(* IEC 61131-3 sources: plc-iiot-stack/flagship/src/POUs/Iiot/FB_IiotKnsMap, 8 files *)

(* ---- ApplyCommand.method.decl.st ---- *)
// Записать принятую команду строки diRule белого списка в GVL_Hmi или GVL_Station (импульс или rValue).
METHOD ApplyCommand : BOOL
VAR_INPUT
    diRule : DINT;
    rValue : REAL;
END_VAR

(* ---- ApplyCommand.method.impl.st ---- *)
ApplyCommand := TRUE;
CASE diRule OF
    1:  // P101 SetAuto
        GVL_Hmi.stP101Cmd.stCommon.xSetAuto := TRUE;
    2:  // P101 SetManual
        GVL_Hmi.stP101Cmd.stCommon.xSetManual := TRUE;
    3:  // P101 Start
        GVL_Hmi.stP101Cmd.xStart := TRUE;
    4:  // P101 Stop
        GVL_Hmi.stP101Cmd.xStop := TRUE;
    5:  // P101 SpeedSp
        GVL_Hmi.stP101Cmd.rSpeedSp_pct := rValue;
    6:  // P101 Ack
        GVL_Hmi.stP101Cmd.stCommon.xAck := TRUE;
    7:  // P101 Reset
        GVL_Hmi.stP101Cmd.stCommon.xReset := TRUE;
    8:  // P102 SetAuto
        GVL_Hmi.stP102Cmd.stCommon.xSetAuto := TRUE;
    9:  // P102 SetManual
        GVL_Hmi.stP102Cmd.stCommon.xSetManual := TRUE;
    10:  // P102 Start
        GVL_Hmi.stP102Cmd.xStart := TRUE;
    11:  // P102 Stop
        GVL_Hmi.stP102Cmd.xStop := TRUE;
    12:  // P102 SpeedSp
        GVL_Hmi.stP102Cmd.rSpeedSp_pct := rValue;
    13:  // P102 Ack
        GVL_Hmi.stP102Cmd.stCommon.xAck := TRUE;
    14:  // P102 Reset
        GVL_Hmi.stP102Cmd.stCommon.xReset := TRUE;
    15:  // P103 SetAuto
        GVL_Hmi.stP103Cmd.stCommon.xSetAuto := TRUE;
    16:  // P103 SetManual
        GVL_Hmi.stP103Cmd.stCommon.xSetManual := TRUE;
    17:  // P103 Start
        GVL_Hmi.stP103Cmd.xStart := TRUE;
    18:  // P103 Stop
        GVL_Hmi.stP103Cmd.xStop := TRUE;
    19:  // P103 SpeedSp
        GVL_Hmi.stP103Cmd.rSpeedSp_pct := rValue;
    20:  // P103 Ack
        GVL_Hmi.stP103Cmd.stCommon.xAck := TRUE;
    21:  // P103 Reset
        GVL_Hmi.stP103Cmd.stCommon.xReset := TRUE;
    22:  // V1 SetAuto
        GVL_Hmi.stV1Cmd.stCommon.xSetAuto := TRUE;
    23:  // V1 SetManual
        GVL_Hmi.stV1Cmd.stCommon.xSetManual := TRUE;
    24:  // V1 Start
        GVL_Hmi.stV1Cmd.xStart := TRUE;
    25:  // V1 Stop
        GVL_Hmi.stV1Cmd.xStop := TRUE;
    26:  // V1 Ack
        GVL_Hmi.stV1Cmd.stCommon.xAck := TRUE;
    27:  // V1 Reset
        GVL_Hmi.stV1Cmd.stCommon.xReset := TRUE;
    28:  // LT101 Ack
        GVL_Hmi.stLT101Cmd.stCommon.xAck := TRUE;
    29:  // LT101 Reset
        GVL_Hmi.stLT101Cmd.stCommon.xReset := TRUE;
    30:  // LS102 Ack
        GVL_Hmi.stLS102Cmd.stCommon.xAck := TRUE;
    31:  // LS102 Reset
        GVL_Hmi.stLS102Cmd.stCommon.xReset := TRUE;
    32:  // LS103 Ack
        GVL_Hmi.stLS103Cmd.stCommon.xAck := TRUE;
    33:  // LS103 Reset
        GVL_Hmi.stLS103Cmd.stCommon.xReset := TRUE;
    34:  // IT111 Ack
        GVL_Hmi.stIT111Cmd.stCommon.xAck := TRUE;
    35:  // IT111 Reset
        GVL_Hmi.stIT111Cmd.stCommon.xReset := TRUE;
    36:  // TS112 Ack
        GVL_Hmi.stTS112Cmd.stCommon.xAck := TRUE;
    37:  // TS112 Reset
        GVL_Hmi.stTS112Cmd.stCommon.xReset := TRUE;
    38:  // MS113 Ack
        GVL_Hmi.stMS113Cmd.stCommon.xAck := TRUE;
    39:  // MS113 Reset
        GVL_Hmi.stMS113Cmd.stCommon.xReset := TRUE;
    40:  // IT121 Ack
        GVL_Hmi.stIT121Cmd.stCommon.xAck := TRUE;
    41:  // IT121 Reset
        GVL_Hmi.stIT121Cmd.stCommon.xReset := TRUE;
    42:  // TS122 Ack
        GVL_Hmi.stTS122Cmd.stCommon.xAck := TRUE;
    43:  // TS122 Reset
        GVL_Hmi.stTS122Cmd.stCommon.xReset := TRUE;
    44:  // MS123 Ack
        GVL_Hmi.stMS123Cmd.stCommon.xAck := TRUE;
    45:  // MS123 Reset
        GVL_Hmi.stMS123Cmd.stCommon.xReset := TRUE;
    46:  // IT131 Ack
        GVL_Hmi.stIT131Cmd.stCommon.xAck := TRUE;
    47:  // IT131 Reset
        GVL_Hmi.stIT131Cmd.stCommon.xReset := TRUE;
    48:  // TS132 Ack
        GVL_Hmi.stTS132Cmd.stCommon.xAck := TRUE;
    49:  // TS132 Reset
        GVL_Hmi.stTS132Cmd.stCommon.xReset := TRUE;
    50:  // MS133 Ack
        GVL_Hmi.stMS133Cmd.stCommon.xAck := TRUE;
    51:  // MS133 Reset
        GVL_Hmi.stMS133Cmd.stCommon.xReset := TRUE;
    52:  // PT201 Ack
        GVL_Hmi.stPT201Cmd.stCommon.xAck := TRUE;
    53:  // PT201 Reset
        GVL_Hmi.stPT201Cmd.stCommon.xReset := TRUE;
    54:  // FT202 Ack
        GVL_Hmi.stFT202Cmd.stCommon.xAck := TRUE;
    55:  // FT202 Reset
        GVL_Hmi.stFT202Cmd.stCommon.xReset := TRUE;
    56:  // LS203 Ack
        GVL_Hmi.stLS203Cmd.stCommon.xAck := TRUE;
    57:  // LS203 Reset
        GVL_Hmi.stLS203Cmd.stCommon.xReset := TRUE;
    58:  // ES301 Ack
        GVL_Hmi.stES301Cmd.stCommon.xAck := TRUE;
    59:  // ES301 Reset
        GVL_Hmi.stES301Cmd.stCommon.xReset := TRUE;
    60:  // YS302 Ack
        GVL_Hmi.stYS302Cmd.stCommon.xAck := TRUE;
    61:  // YS302 Reset
        GVL_Hmi.stYS302Cmd.stCommon.xReset := TRUE;
    62:  // YS303 Ack
        GVL_Hmi.stYS303Cmd.stCommon.xAck := TRUE;
    63:  // YS303 Reset
        GVL_Hmi.stYS303Cmd.stCommon.xReset := TRUE;
    64:  // AT401 Ack
        GVL_Hmi.stAT401Cmd.stCommon.xAck := TRUE;
    65:  // AT401 Reset
        GVL_Hmi.stAT401Cmd.stCommon.xReset := TRUE;
    66:  // AT402 Ack
        GVL_Hmi.stAT402Cmd.stCommon.xAck := TRUE;
    67:  // AT402 Reset
        GVL_Hmi.stAT402Cmd.stCommon.xReset := TRUE;
    68:  // TT403 Ack
        GVL_Hmi.stTT403Cmd.stCommon.xAck := TRUE;
    69:  // TT403 Reset
        GVL_Hmi.stTT403Cmd.stCommon.xReset := TRUE;
    70:  // ZS404 Ack
        GVL_Hmi.stZS404Cmd.stCommon.xAck := TRUE;
    71:  // ZS404 Reset
        GVL_Hmi.stZS404Cmd.stCommon.xReset := TRUE;
    72:  // YS405 Ack
        GVL_Hmi.stYS405Cmd.stCommon.xAck := TRUE;
    73:  // YS405 Reset
        GVL_Hmi.stYS405Cmd.stCommon.xReset := TRUE;
    74:  // HS501 Ack
        GVL_Hmi.stHS501Cmd.stCommon.xAck := TRUE;
    75:  // HS501 Reset
        GVL_Hmi.stHS501Cmd.stCommon.xReset := TRUE;
    76:  // HS502 Ack
        GVL_Hmi.stHS502Cmd.stCommon.xAck := TRUE;
    77:  // HS502 Reset
        GVL_Hmi.stHS502Cmd.stCommon.xReset := TRUE;
    78:  // KNS1 SetAuto
        GVL_Station.stStationCmd.xSetAuto := TRUE;
    79:  // KNS1 SetManual
        GVL_Station.stStationCmd.xSetManual := TRUE;
    80:  // KNS1 SetStepped
        GVL_Station.stStationCmd.xSetStepped := TRUE;
    81:  // KNS1 SetLevelPid
        GVL_Station.stStationCmd.xSetLevelPid := TRUE;
    82:  // KNS1 AckAll
        GVL_Station.stStationCmd.xAckAll := TRUE;
    83:  // KNS1 ResetAll
        GVL_Station.stStationCmd.xResetAll := TRUE;
    84:  // KNS1 Silence
        GVL_Station.stStationCmd.xSilence := TRUE;
    85:  // LIC101 SetAuto
        GVL_Station.stLIC101Cmd.stCommon.xSetAuto := TRUE;
    86:  // LIC101 SetManual
        GVL_Station.stLIC101Cmd.stCommon.xSetManual := TRUE;
ELSE
    ApplyCommand := FALSE;
END_CASE

(* ---- DeviceCmdState.method.decl.st ---- *)
// Счётчик обработанных команд и результат последней команды устройства diDev (ST_IiotCmdRule.diDev).
METHOD DeviceCmdState
VAR_INPUT
    diDev : DINT;
END_VAR
VAR_OUTPUT
    uiSeq : UINT;
    iResult : INT;
END_VAR

(* ---- DeviceCmdState.method.impl.st ---- *)
uiSeq := 0;
iResult := 0;
CASE diDev OF
    1:  // P101
        uiSeq := GVL_Devices.fbP101.stSts.stCommon.uiCmdSeq;
        iResult := TO_INT(GVL_Devices.fbP101.stSts.stCommon.eCmdResult);
    2:  // P102
        uiSeq := GVL_Devices.fbP102.stSts.stCommon.uiCmdSeq;
        iResult := TO_INT(GVL_Devices.fbP102.stSts.stCommon.eCmdResult);
    3:  // P103
        uiSeq := GVL_Devices.fbP103.stSts.stCommon.uiCmdSeq;
        iResult := TO_INT(GVL_Devices.fbP103.stSts.stCommon.eCmdResult);
    4:  // V1
        uiSeq := GVL_Devices.fbV1.stSts.stCommon.uiCmdSeq;
        iResult := TO_INT(GVL_Devices.fbV1.stSts.stCommon.eCmdResult);
    5:  // LT101
        uiSeq := GVL_Devices.fbLT101.stSts.stCommon.uiCmdSeq;
        iResult := TO_INT(GVL_Devices.fbLT101.stSts.stCommon.eCmdResult);
    6:  // LS102
        uiSeq := GVL_Devices.fbLS102.stSts.stCommon.uiCmdSeq;
        iResult := TO_INT(GVL_Devices.fbLS102.stSts.stCommon.eCmdResult);
    7:  // LS103
        uiSeq := GVL_Devices.fbLS103.stSts.stCommon.uiCmdSeq;
        iResult := TO_INT(GVL_Devices.fbLS103.stSts.stCommon.eCmdResult);
    8:  // IT111
        uiSeq := GVL_Devices.fbIT111.stSts.stCommon.uiCmdSeq;
        iResult := TO_INT(GVL_Devices.fbIT111.stSts.stCommon.eCmdResult);
    9:  // TS112
        uiSeq := GVL_Devices.fbTS112.stSts.stCommon.uiCmdSeq;
        iResult := TO_INT(GVL_Devices.fbTS112.stSts.stCommon.eCmdResult);
    10:  // MS113
        uiSeq := GVL_Devices.fbMS113.stSts.stCommon.uiCmdSeq;
        iResult := TO_INT(GVL_Devices.fbMS113.stSts.stCommon.eCmdResult);
    11:  // IT121
        uiSeq := GVL_Devices.fbIT121.stSts.stCommon.uiCmdSeq;
        iResult := TO_INT(GVL_Devices.fbIT121.stSts.stCommon.eCmdResult);
    12:  // TS122
        uiSeq := GVL_Devices.fbTS122.stSts.stCommon.uiCmdSeq;
        iResult := TO_INT(GVL_Devices.fbTS122.stSts.stCommon.eCmdResult);
    13:  // MS123
        uiSeq := GVL_Devices.fbMS123.stSts.stCommon.uiCmdSeq;
        iResult := TO_INT(GVL_Devices.fbMS123.stSts.stCommon.eCmdResult);
    14:  // IT131
        uiSeq := GVL_Devices.fbIT131.stSts.stCommon.uiCmdSeq;
        iResult := TO_INT(GVL_Devices.fbIT131.stSts.stCommon.eCmdResult);
    15:  // TS132
        uiSeq := GVL_Devices.fbTS132.stSts.stCommon.uiCmdSeq;
        iResult := TO_INT(GVL_Devices.fbTS132.stSts.stCommon.eCmdResult);
    16:  // MS133
        uiSeq := GVL_Devices.fbMS133.stSts.stCommon.uiCmdSeq;
        iResult := TO_INT(GVL_Devices.fbMS133.stSts.stCommon.eCmdResult);
    17:  // PT201
        uiSeq := GVL_Devices.fbPT201.stSts.stCommon.uiCmdSeq;
        iResult := TO_INT(GVL_Devices.fbPT201.stSts.stCommon.eCmdResult);
    18:  // FT202
        uiSeq := GVL_Devices.fbFT202.stSts.stCommon.uiCmdSeq;
        iResult := TO_INT(GVL_Devices.fbFT202.stSts.stCommon.eCmdResult);
    19:  // LS203
        uiSeq := GVL_Devices.fbLS203.stSts.stCommon.uiCmdSeq;
        iResult := TO_INT(GVL_Devices.fbLS203.stSts.stCommon.eCmdResult);
    20:  // ES301
        uiSeq := GVL_Devices.fbES301.stSts.stCommon.uiCmdSeq;
        iResult := TO_INT(GVL_Devices.fbES301.stSts.stCommon.eCmdResult);
    21:  // YS302
        uiSeq := GVL_Devices.fbYS302.stSts.stCommon.uiCmdSeq;
        iResult := TO_INT(GVL_Devices.fbYS302.stSts.stCommon.eCmdResult);
    22:  // YS303
        uiSeq := GVL_Devices.fbYS303.stSts.stCommon.uiCmdSeq;
        iResult := TO_INT(GVL_Devices.fbYS303.stSts.stCommon.eCmdResult);
    23:  // AT401
        uiSeq := GVL_Devices.fbAT401.stSts.stCommon.uiCmdSeq;
        iResult := TO_INT(GVL_Devices.fbAT401.stSts.stCommon.eCmdResult);
    24:  // AT402
        uiSeq := GVL_Devices.fbAT402.stSts.stCommon.uiCmdSeq;
        iResult := TO_INT(GVL_Devices.fbAT402.stSts.stCommon.eCmdResult);
    25:  // TT403
        uiSeq := GVL_Devices.fbTT403.stSts.stCommon.uiCmdSeq;
        iResult := TO_INT(GVL_Devices.fbTT403.stSts.stCommon.eCmdResult);
    26:  // ZS404
        uiSeq := GVL_Devices.fbZS404.stSts.stCommon.uiCmdSeq;
        iResult := TO_INT(GVL_Devices.fbZS404.stSts.stCommon.eCmdResult);
    27:  // YS405
        uiSeq := GVL_Devices.fbYS405.stSts.stCommon.uiCmdSeq;
        iResult := TO_INT(GVL_Devices.fbYS405.stSts.stCommon.eCmdResult);
    28:  // HS501
        uiSeq := GVL_Devices.fbHS501.stSts.stCommon.uiCmdSeq;
        iResult := TO_INT(GVL_Devices.fbHS501.stSts.stCommon.eCmdResult);
    29:  // HS502
        uiSeq := GVL_Devices.fbHS502.stSts.stCommon.uiCmdSeq;
        iResult := TO_INT(GVL_Devices.fbHS502.stSts.stCommon.eCmdResult);
    30:  // KNS1
        uiSeq := GVL_Station.stStationSts.uiCmdSeq;
        iResult := TO_INT(GVL_Station.stStationSts.eCmdResult);
    31:  // LIC101
        uiSeq := GVL_Station.fbLIC101.stSts.stCommon.uiCmdSeq;
        iResult := TO_INT(GVL_Station.fbLIC101.stSts.stCommon.eCmdResult);
END_CASE

(* ---- FillAlarmWords.method.decl.st ---- *)
// Слова тревог устройств и станции (строки — источники перечня тревог по порядку ALARM_CFG.diWords).
METHOD FillAlarmWords
VAR_IN_OUT
    aWordTable : ARRAY[*] OF ST_IiotAlarmWords;
END_VAR

(* ---- FillAlarmWords.method.impl.st ---- *)
// Массив меньше перечня (не тот, что объявлен в PRG_Iiot): ничего не пишем, а не выходим за границы
IF LOWER_BOUND(aWordTable, 1) > 1 OR UPPER_BOUND(aWordTable, 1) < GVL_IiotMap.ALARM_WORDS_COUNT THEN
    RETURN;
END_IF
aWordTable[1].wActive := GVL_Devices.fbP101.stSts.stCommon.wAlmActive;
aWordTable[1].wUnack := GVL_Devices.fbP101.stSts.stCommon.wAlmUnack;
aWordTable[1].wShelved := GVL_Devices.fbP101.stSts.stCommon.wAlmShelved;
aWordTable[1].wSuppressed := GVL_Devices.fbP101.stSts.stCommon.wAlmSuppressed;
aWordTable[1].xOutOfService := GVL_Devices.fbP101.stSts.stCommon.eMode = PL.E_DeviceMode.OutOfService;
aWordTable[2].wActive := GVL_Devices.fbP102.stSts.stCommon.wAlmActive;
aWordTable[2].wUnack := GVL_Devices.fbP102.stSts.stCommon.wAlmUnack;
aWordTable[2].wShelved := GVL_Devices.fbP102.stSts.stCommon.wAlmShelved;
aWordTable[2].wSuppressed := GVL_Devices.fbP102.stSts.stCommon.wAlmSuppressed;
aWordTable[2].xOutOfService := GVL_Devices.fbP102.stSts.stCommon.eMode = PL.E_DeviceMode.OutOfService;
aWordTable[3].wActive := GVL_Devices.fbP103.stSts.stCommon.wAlmActive;
aWordTable[3].wUnack := GVL_Devices.fbP103.stSts.stCommon.wAlmUnack;
aWordTable[3].wShelved := GVL_Devices.fbP103.stSts.stCommon.wAlmShelved;
aWordTable[3].wSuppressed := GVL_Devices.fbP103.stSts.stCommon.wAlmSuppressed;
aWordTable[3].xOutOfService := GVL_Devices.fbP103.stSts.stCommon.eMode = PL.E_DeviceMode.OutOfService;
aWordTable[4].wActive := GVL_Devices.fbV1.stSts.stCommon.wAlmActive;
aWordTable[4].wUnack := GVL_Devices.fbV1.stSts.stCommon.wAlmUnack;
aWordTable[4].wShelved := GVL_Devices.fbV1.stSts.stCommon.wAlmShelved;
aWordTable[4].wSuppressed := GVL_Devices.fbV1.stSts.stCommon.wAlmSuppressed;
aWordTable[4].xOutOfService := GVL_Devices.fbV1.stSts.stCommon.eMode = PL.E_DeviceMode.OutOfService;
aWordTable[5].wActive := GVL_Devices.fbLT101.stSts.stCommon.wAlmActive;
aWordTable[5].wUnack := GVL_Devices.fbLT101.stSts.stCommon.wAlmUnack;
aWordTable[5].wShelved := GVL_Devices.fbLT101.stSts.stCommon.wAlmShelved;
aWordTable[5].wSuppressed := GVL_Devices.fbLT101.stSts.stCommon.wAlmSuppressed;
aWordTable[5].xOutOfService := GVL_Devices.fbLT101.stSts.stCommon.eMode = PL.E_DeviceMode.OutOfService;
aWordTable[6].wActive := GVL_Devices.fbLS102.stSts.stCommon.wAlmActive;
aWordTable[6].wUnack := GVL_Devices.fbLS102.stSts.stCommon.wAlmUnack;
aWordTable[6].wShelved := GVL_Devices.fbLS102.stSts.stCommon.wAlmShelved;
aWordTable[6].wSuppressed := GVL_Devices.fbLS102.stSts.stCommon.wAlmSuppressed;
aWordTable[6].xOutOfService := GVL_Devices.fbLS102.stSts.stCommon.eMode = PL.E_DeviceMode.OutOfService;
aWordTable[7].wActive := GVL_Devices.fbLS103.stSts.stCommon.wAlmActive;
aWordTable[7].wUnack := GVL_Devices.fbLS103.stSts.stCommon.wAlmUnack;
aWordTable[7].wShelved := GVL_Devices.fbLS103.stSts.stCommon.wAlmShelved;
aWordTable[7].wSuppressed := GVL_Devices.fbLS103.stSts.stCommon.wAlmSuppressed;
aWordTable[7].xOutOfService := GVL_Devices.fbLS103.stSts.stCommon.eMode = PL.E_DeviceMode.OutOfService;
aWordTable[8].wActive := GVL_Devices.fbIT111.stSts.stCommon.wAlmActive;
aWordTable[8].wUnack := GVL_Devices.fbIT111.stSts.stCommon.wAlmUnack;
aWordTable[8].wShelved := GVL_Devices.fbIT111.stSts.stCommon.wAlmShelved;
aWordTable[8].wSuppressed := GVL_Devices.fbIT111.stSts.stCommon.wAlmSuppressed;
aWordTable[8].xOutOfService := GVL_Devices.fbIT111.stSts.stCommon.eMode = PL.E_DeviceMode.OutOfService;
aWordTable[9].wActive := GVL_Devices.fbTS112.stSts.stCommon.wAlmActive;
aWordTable[9].wUnack := GVL_Devices.fbTS112.stSts.stCommon.wAlmUnack;
aWordTable[9].wShelved := GVL_Devices.fbTS112.stSts.stCommon.wAlmShelved;
aWordTable[9].wSuppressed := GVL_Devices.fbTS112.stSts.stCommon.wAlmSuppressed;
aWordTable[9].xOutOfService := GVL_Devices.fbTS112.stSts.stCommon.eMode = PL.E_DeviceMode.OutOfService;
aWordTable[10].wActive := GVL_Devices.fbMS113.stSts.stCommon.wAlmActive;
aWordTable[10].wUnack := GVL_Devices.fbMS113.stSts.stCommon.wAlmUnack;
aWordTable[10].wShelved := GVL_Devices.fbMS113.stSts.stCommon.wAlmShelved;
aWordTable[10].wSuppressed := GVL_Devices.fbMS113.stSts.stCommon.wAlmSuppressed;
aWordTable[10].xOutOfService := GVL_Devices.fbMS113.stSts.stCommon.eMode = PL.E_DeviceMode.OutOfService;
aWordTable[11].wActive := GVL_Devices.fbIT121.stSts.stCommon.wAlmActive;
aWordTable[11].wUnack := GVL_Devices.fbIT121.stSts.stCommon.wAlmUnack;
aWordTable[11].wShelved := GVL_Devices.fbIT121.stSts.stCommon.wAlmShelved;
aWordTable[11].wSuppressed := GVL_Devices.fbIT121.stSts.stCommon.wAlmSuppressed;
aWordTable[11].xOutOfService := GVL_Devices.fbIT121.stSts.stCommon.eMode = PL.E_DeviceMode.OutOfService;
aWordTable[12].wActive := GVL_Devices.fbTS122.stSts.stCommon.wAlmActive;
aWordTable[12].wUnack := GVL_Devices.fbTS122.stSts.stCommon.wAlmUnack;
aWordTable[12].wShelved := GVL_Devices.fbTS122.stSts.stCommon.wAlmShelved;
aWordTable[12].wSuppressed := GVL_Devices.fbTS122.stSts.stCommon.wAlmSuppressed;
aWordTable[12].xOutOfService := GVL_Devices.fbTS122.stSts.stCommon.eMode = PL.E_DeviceMode.OutOfService;
aWordTable[13].wActive := GVL_Devices.fbMS123.stSts.stCommon.wAlmActive;
aWordTable[13].wUnack := GVL_Devices.fbMS123.stSts.stCommon.wAlmUnack;
aWordTable[13].wShelved := GVL_Devices.fbMS123.stSts.stCommon.wAlmShelved;
aWordTable[13].wSuppressed := GVL_Devices.fbMS123.stSts.stCommon.wAlmSuppressed;
aWordTable[13].xOutOfService := GVL_Devices.fbMS123.stSts.stCommon.eMode = PL.E_DeviceMode.OutOfService;
aWordTable[14].wActive := GVL_Devices.fbIT131.stSts.stCommon.wAlmActive;
aWordTable[14].wUnack := GVL_Devices.fbIT131.stSts.stCommon.wAlmUnack;
aWordTable[14].wShelved := GVL_Devices.fbIT131.stSts.stCommon.wAlmShelved;
aWordTable[14].wSuppressed := GVL_Devices.fbIT131.stSts.stCommon.wAlmSuppressed;
aWordTable[14].xOutOfService := GVL_Devices.fbIT131.stSts.stCommon.eMode = PL.E_DeviceMode.OutOfService;
aWordTable[15].wActive := GVL_Devices.fbTS132.stSts.stCommon.wAlmActive;
aWordTable[15].wUnack := GVL_Devices.fbTS132.stSts.stCommon.wAlmUnack;
aWordTable[15].wShelved := GVL_Devices.fbTS132.stSts.stCommon.wAlmShelved;
aWordTable[15].wSuppressed := GVL_Devices.fbTS132.stSts.stCommon.wAlmSuppressed;
aWordTable[15].xOutOfService := GVL_Devices.fbTS132.stSts.stCommon.eMode = PL.E_DeviceMode.OutOfService;
aWordTable[16].wActive := GVL_Devices.fbMS133.stSts.stCommon.wAlmActive;
aWordTable[16].wUnack := GVL_Devices.fbMS133.stSts.stCommon.wAlmUnack;
aWordTable[16].wShelved := GVL_Devices.fbMS133.stSts.stCommon.wAlmShelved;
aWordTable[16].wSuppressed := GVL_Devices.fbMS133.stSts.stCommon.wAlmSuppressed;
aWordTable[16].xOutOfService := GVL_Devices.fbMS133.stSts.stCommon.eMode = PL.E_DeviceMode.OutOfService;
aWordTable[17].wActive := GVL_Devices.fbPT201.stSts.stCommon.wAlmActive;
aWordTable[17].wUnack := GVL_Devices.fbPT201.stSts.stCommon.wAlmUnack;
aWordTable[17].wShelved := GVL_Devices.fbPT201.stSts.stCommon.wAlmShelved;
aWordTable[17].wSuppressed := GVL_Devices.fbPT201.stSts.stCommon.wAlmSuppressed;
aWordTable[17].xOutOfService := GVL_Devices.fbPT201.stSts.stCommon.eMode = PL.E_DeviceMode.OutOfService;
aWordTable[18].wActive := GVL_Devices.fbFT202.stSts.stCommon.wAlmActive;
aWordTable[18].wUnack := GVL_Devices.fbFT202.stSts.stCommon.wAlmUnack;
aWordTable[18].wShelved := GVL_Devices.fbFT202.stSts.stCommon.wAlmShelved;
aWordTable[18].wSuppressed := GVL_Devices.fbFT202.stSts.stCommon.wAlmSuppressed;
aWordTable[18].xOutOfService := GVL_Devices.fbFT202.stSts.stCommon.eMode = PL.E_DeviceMode.OutOfService;
aWordTable[19].wActive := GVL_Devices.fbLS203.stSts.stCommon.wAlmActive;
aWordTable[19].wUnack := GVL_Devices.fbLS203.stSts.stCommon.wAlmUnack;
aWordTable[19].wShelved := GVL_Devices.fbLS203.stSts.stCommon.wAlmShelved;
aWordTable[19].wSuppressed := GVL_Devices.fbLS203.stSts.stCommon.wAlmSuppressed;
aWordTable[19].xOutOfService := GVL_Devices.fbLS203.stSts.stCommon.eMode = PL.E_DeviceMode.OutOfService;
aWordTable[20].wActive := GVL_Devices.fbES301.stSts.stCommon.wAlmActive;
aWordTable[20].wUnack := GVL_Devices.fbES301.stSts.stCommon.wAlmUnack;
aWordTable[20].wShelved := GVL_Devices.fbES301.stSts.stCommon.wAlmShelved;
aWordTable[20].wSuppressed := GVL_Devices.fbES301.stSts.stCommon.wAlmSuppressed;
aWordTable[20].xOutOfService := GVL_Devices.fbES301.stSts.stCommon.eMode = PL.E_DeviceMode.OutOfService;
aWordTable[21].wActive := GVL_Devices.fbYS302.stSts.stCommon.wAlmActive;
aWordTable[21].wUnack := GVL_Devices.fbYS302.stSts.stCommon.wAlmUnack;
aWordTable[21].wShelved := GVL_Devices.fbYS302.stSts.stCommon.wAlmShelved;
aWordTable[21].wSuppressed := GVL_Devices.fbYS302.stSts.stCommon.wAlmSuppressed;
aWordTable[21].xOutOfService := GVL_Devices.fbYS302.stSts.stCommon.eMode = PL.E_DeviceMode.OutOfService;
aWordTable[22].wActive := GVL_Devices.fbYS303.stSts.stCommon.wAlmActive;
aWordTable[22].wUnack := GVL_Devices.fbYS303.stSts.stCommon.wAlmUnack;
aWordTable[22].wShelved := GVL_Devices.fbYS303.stSts.stCommon.wAlmShelved;
aWordTable[22].wSuppressed := GVL_Devices.fbYS303.stSts.stCommon.wAlmSuppressed;
aWordTable[22].xOutOfService := GVL_Devices.fbYS303.stSts.stCommon.eMode = PL.E_DeviceMode.OutOfService;
aWordTable[23].wActive := GVL_Devices.fbAT401.stSts.stCommon.wAlmActive;
aWordTable[23].wUnack := GVL_Devices.fbAT401.stSts.stCommon.wAlmUnack;
aWordTable[23].wShelved := GVL_Devices.fbAT401.stSts.stCommon.wAlmShelved;
aWordTable[23].wSuppressed := GVL_Devices.fbAT401.stSts.stCommon.wAlmSuppressed;
aWordTable[23].xOutOfService := GVL_Devices.fbAT401.stSts.stCommon.eMode = PL.E_DeviceMode.OutOfService;
aWordTable[24].wActive := GVL_Devices.fbAT402.stSts.stCommon.wAlmActive;
aWordTable[24].wUnack := GVL_Devices.fbAT402.stSts.stCommon.wAlmUnack;
aWordTable[24].wShelved := GVL_Devices.fbAT402.stSts.stCommon.wAlmShelved;
aWordTable[24].wSuppressed := GVL_Devices.fbAT402.stSts.stCommon.wAlmSuppressed;
aWordTable[24].xOutOfService := GVL_Devices.fbAT402.stSts.stCommon.eMode = PL.E_DeviceMode.OutOfService;
aWordTable[25].wActive := GVL_Devices.fbTT403.stSts.stCommon.wAlmActive;
aWordTable[25].wUnack := GVL_Devices.fbTT403.stSts.stCommon.wAlmUnack;
aWordTable[25].wShelved := GVL_Devices.fbTT403.stSts.stCommon.wAlmShelved;
aWordTable[25].wSuppressed := GVL_Devices.fbTT403.stSts.stCommon.wAlmSuppressed;
aWordTable[25].xOutOfService := GVL_Devices.fbTT403.stSts.stCommon.eMode = PL.E_DeviceMode.OutOfService;
aWordTable[26].wActive := GVL_Devices.fbZS404.stSts.stCommon.wAlmActive;
aWordTable[26].wUnack := GVL_Devices.fbZS404.stSts.stCommon.wAlmUnack;
aWordTable[26].wShelved := GVL_Devices.fbZS404.stSts.stCommon.wAlmShelved;
aWordTable[26].wSuppressed := GVL_Devices.fbZS404.stSts.stCommon.wAlmSuppressed;
aWordTable[26].xOutOfService := GVL_Devices.fbZS404.stSts.stCommon.eMode = PL.E_DeviceMode.OutOfService;
aWordTable[27].wActive := GVL_Devices.fbYS405.stSts.stCommon.wAlmActive;
aWordTable[27].wUnack := GVL_Devices.fbYS405.stSts.stCommon.wAlmUnack;
aWordTable[27].wShelved := GVL_Devices.fbYS405.stSts.stCommon.wAlmShelved;
aWordTable[27].wSuppressed := GVL_Devices.fbYS405.stSts.stCommon.wAlmSuppressed;
aWordTable[27].xOutOfService := GVL_Devices.fbYS405.stSts.stCommon.eMode = PL.E_DeviceMode.OutOfService;
aWordTable[28].wActive := GVL_Station.stStationSts.wAlmActive;
aWordTable[28].wUnack := GVL_Station.stStationSts.wAlmUnack;
aWordTable[28].wShelved := GVL_Station.stStationSts.wAlmShelved;
aWordTable[28].wSuppressed := 0;
aWordTable[28].xOutOfService := FALSE;

(* ---- FillPoints.method.decl.st ---- *)
// Значения и качество метрик с путём в ПЛК (метрики узла PLC1 заполняет PRG_Iiot).
METHOD FillPoints
VAR_IN_OUT
    aPointTable : ARRAY[*] OF ST_IiotPoint;
END_VAR

(* ---- FillPoints.method.impl.st ---- *)
// Массив меньше перечня (не тот, что объявлен в PRG_Iiot): ничего не пишем, а не выходим за границы
IF LOWER_BOUND(aPointTable, 1) > 1 OR UPPER_BOUND(aPointTable, 1) < GVL_IiotMap.POINT_COUNT THEN
    RETURN;
END_IF
aPointTable[1].lrValue := BOOL_TO_LREAL(GVL_Devices.fbP101.xRunning);
aPointTable[1].eQuality := F_IiotQuality(xValid := TRUE, iNe107 := TO_INT(GVL_Devices.fbP101.stSts.stCommon.eNe107));
aPointTable[2].lrValue := INT_TO_LREAL(TO_INT(GVL_Devices.fbP101.stSts.eState));
aPointTable[2].eQuality := F_IiotQuality(xValid := TRUE, iNe107 := TO_INT(GVL_Devices.fbP101.stSts.stCommon.eNe107));
aPointTable[3].lrValue := REAL_TO_LREAL(GVL_Devices.fbP101.stSts.rSpeedAct_pct);
aPointTable[3].eQuality := F_IiotQuality(xValid := TRUE, iNe107 := TO_INT(GVL_Devices.fbP101.stSts.stCommon.eNe107));
IF (GVL_Devices.fbP101.stSts.stCommon.wFault AND PL.GVL_Const.MOT_FLT_COMM_LOSS) <> 0
   OR (GVL_Devices.fbP101.stSts.stCommon.wWarning AND PL.GVL_Const.MOT_WRN_COMM_LOSS) <> 0 THEN
    aPointTable[3].eQuality := E_IiotQuality.Bad;
END_IF
aPointTable[4].lrValue := REAL_TO_LREAL(GVL_Devices.fbP101.stSts.rSpeedRef_pct);
aPointTable[4].eQuality := F_IiotQuality(xValid := TRUE, iNe107 := TO_INT(GVL_Devices.fbP101.stSts.stCommon.eNe107));
aPointTable[5].lrValue := REAL_TO_LREAL(GVL_Devices.fbP101.stSts.rRunTime_h);
aPointTable[5].eQuality := F_IiotQuality(xValid := TRUE, iNe107 := TO_INT(GVL_Devices.fbP101.stSts.stCommon.eNe107));
aPointTable[6].lrValue := UDINT_TO_LREAL(GVL_Devices.fbP101.stSts.udiStarts);
aPointTable[6].eQuality := F_IiotQuality(xValid := TRUE, iNe107 := TO_INT(GVL_Devices.fbP101.stSts.stCommon.eNe107));
aPointTable[7].lrValue := UINT_TO_LREAL(GVL_Devices.fbP101.stSts.uiStartsLastHour);
aPointTable[7].eQuality := F_IiotQuality(xValid := TRUE, iNe107 := TO_INT(GVL_Devices.fbP101.stSts.stCommon.eNe107));
aPointTable[8].lrValue := REAL_TO_LREAL(GVL_Devices.fbP101.stSts.rRunTimeMaint_h);
aPointTable[8].eQuality := F_IiotQuality(xValid := TRUE, iNe107 := TO_INT(GVL_Devices.fbP101.stSts.stCommon.eNe107));
aPointTable[9].lrValue := UDINT_TO_LREAL(GVL_Devices.fbP101.stSts.udiStartsMaint);
aPointTable[9].eQuality := F_IiotQuality(xValid := TRUE, iNe107 := TO_INT(GVL_Devices.fbP101.stSts.stCommon.eNe107));
aPointTable[10].lrValue := UINT_TO_LREAL(GVL_IO.uiP101_FCODE);
aPointTable[10].eQuality := F_IiotQuality(xValid := TRUE, iNe107 := TO_INT(GVL_Devices.fbP101.stSts.stCommon.eNe107));
IF (GVL_Devices.fbP101.stSts.stCommon.wFault AND PL.GVL_Const.MOT_FLT_COMM_LOSS) <> 0
   OR (GVL_Devices.fbP101.stSts.stCommon.wWarning AND PL.GVL_Const.MOT_WRN_COMM_LOSS) <> 0 THEN
    aPointTable[10].eQuality := E_IiotQuality.Bad;
END_IF
aPointTable[11].lrValue := INT_TO_LREAL(TO_INT(GVL_Devices.fbP101.stSts.stCommon.eMode));
aPointTable[11].eQuality := F_IiotQuality(xValid := TRUE, iNe107 := TO_INT(GVL_Devices.fbP101.stSts.stCommon.eNe107));
aPointTable[12].lrValue := INT_TO_LREAL(TO_INT(GVL_Devices.fbP101.stSts.stCommon.eNe107));
aPointTable[12].eQuality := F_IiotQuality(xValid := TRUE, iNe107 := TO_INT(GVL_Devices.fbP101.stSts.stCommon.eNe107));
aPointTable[13].lrValue := BOOL_TO_LREAL(GVL_Devices.fbP102.xRunning);
aPointTable[13].eQuality := F_IiotQuality(xValid := TRUE, iNe107 := TO_INT(GVL_Devices.fbP102.stSts.stCommon.eNe107));
aPointTable[14].lrValue := INT_TO_LREAL(TO_INT(GVL_Devices.fbP102.stSts.eState));
aPointTable[14].eQuality := F_IiotQuality(xValid := TRUE, iNe107 := TO_INT(GVL_Devices.fbP102.stSts.stCommon.eNe107));
aPointTable[15].lrValue := REAL_TO_LREAL(GVL_Devices.fbP102.stSts.rSpeedAct_pct);
aPointTable[15].eQuality := F_IiotQuality(xValid := TRUE, iNe107 := TO_INT(GVL_Devices.fbP102.stSts.stCommon.eNe107));
IF (GVL_Devices.fbP102.stSts.stCommon.wFault AND PL.GVL_Const.MOT_FLT_COMM_LOSS) <> 0
   OR (GVL_Devices.fbP102.stSts.stCommon.wWarning AND PL.GVL_Const.MOT_WRN_COMM_LOSS) <> 0 THEN
    aPointTable[15].eQuality := E_IiotQuality.Bad;
END_IF
aPointTable[16].lrValue := REAL_TO_LREAL(GVL_Devices.fbP102.stSts.rSpeedRef_pct);
aPointTable[16].eQuality := F_IiotQuality(xValid := TRUE, iNe107 := TO_INT(GVL_Devices.fbP102.stSts.stCommon.eNe107));
aPointTable[17].lrValue := REAL_TO_LREAL(GVL_Devices.fbP102.stSts.rRunTime_h);
aPointTable[17].eQuality := F_IiotQuality(xValid := TRUE, iNe107 := TO_INT(GVL_Devices.fbP102.stSts.stCommon.eNe107));
aPointTable[18].lrValue := UDINT_TO_LREAL(GVL_Devices.fbP102.stSts.udiStarts);
aPointTable[18].eQuality := F_IiotQuality(xValid := TRUE, iNe107 := TO_INT(GVL_Devices.fbP102.stSts.stCommon.eNe107));
aPointTable[19].lrValue := UINT_TO_LREAL(GVL_Devices.fbP102.stSts.uiStartsLastHour);
aPointTable[19].eQuality := F_IiotQuality(xValid := TRUE, iNe107 := TO_INT(GVL_Devices.fbP102.stSts.stCommon.eNe107));
aPointTable[20].lrValue := REAL_TO_LREAL(GVL_Devices.fbP102.stSts.rRunTimeMaint_h);
aPointTable[20].eQuality := F_IiotQuality(xValid := TRUE, iNe107 := TO_INT(GVL_Devices.fbP102.stSts.stCommon.eNe107));
aPointTable[21].lrValue := UDINT_TO_LREAL(GVL_Devices.fbP102.stSts.udiStartsMaint);
aPointTable[21].eQuality := F_IiotQuality(xValid := TRUE, iNe107 := TO_INT(GVL_Devices.fbP102.stSts.stCommon.eNe107));
aPointTable[22].lrValue := UINT_TO_LREAL(GVL_IO.uiP102_FCODE);
aPointTable[22].eQuality := F_IiotQuality(xValid := TRUE, iNe107 := TO_INT(GVL_Devices.fbP102.stSts.stCommon.eNe107));
IF (GVL_Devices.fbP102.stSts.stCommon.wFault AND PL.GVL_Const.MOT_FLT_COMM_LOSS) <> 0
   OR (GVL_Devices.fbP102.stSts.stCommon.wWarning AND PL.GVL_Const.MOT_WRN_COMM_LOSS) <> 0 THEN
    aPointTable[22].eQuality := E_IiotQuality.Bad;
END_IF
aPointTable[23].lrValue := INT_TO_LREAL(TO_INT(GVL_Devices.fbP102.stSts.stCommon.eMode));
aPointTable[23].eQuality := F_IiotQuality(xValid := TRUE, iNe107 := TO_INT(GVL_Devices.fbP102.stSts.stCommon.eNe107));
aPointTable[24].lrValue := INT_TO_LREAL(TO_INT(GVL_Devices.fbP102.stSts.stCommon.eNe107));
aPointTable[24].eQuality := F_IiotQuality(xValid := TRUE, iNe107 := TO_INT(GVL_Devices.fbP102.stSts.stCommon.eNe107));
aPointTable[25].lrValue := BOOL_TO_LREAL(GVL_Devices.fbP103.xRunning);
aPointTable[25].eQuality := F_IiotQuality(xValid := TRUE, iNe107 := TO_INT(GVL_Devices.fbP103.stSts.stCommon.eNe107));
aPointTable[26].lrValue := INT_TO_LREAL(TO_INT(GVL_Devices.fbP103.stSts.eState));
aPointTable[26].eQuality := F_IiotQuality(xValid := TRUE, iNe107 := TO_INT(GVL_Devices.fbP103.stSts.stCommon.eNe107));
aPointTable[27].lrValue := REAL_TO_LREAL(GVL_Devices.fbP103.stSts.rSpeedAct_pct);
aPointTable[27].eQuality := F_IiotQuality(xValid := TRUE, iNe107 := TO_INT(GVL_Devices.fbP103.stSts.stCommon.eNe107));
IF (GVL_Devices.fbP103.stSts.stCommon.wFault AND PL.GVL_Const.MOT_FLT_COMM_LOSS) <> 0
   OR (GVL_Devices.fbP103.stSts.stCommon.wWarning AND PL.GVL_Const.MOT_WRN_COMM_LOSS) <> 0 THEN
    aPointTable[27].eQuality := E_IiotQuality.Bad;
END_IF
aPointTable[28].lrValue := REAL_TO_LREAL(GVL_Devices.fbP103.stSts.rSpeedRef_pct);
aPointTable[28].eQuality := F_IiotQuality(xValid := TRUE, iNe107 := TO_INT(GVL_Devices.fbP103.stSts.stCommon.eNe107));
aPointTable[29].lrValue := REAL_TO_LREAL(GVL_Devices.fbP103.stSts.rRunTime_h);
aPointTable[29].eQuality := F_IiotQuality(xValid := TRUE, iNe107 := TO_INT(GVL_Devices.fbP103.stSts.stCommon.eNe107));
aPointTable[30].lrValue := UDINT_TO_LREAL(GVL_Devices.fbP103.stSts.udiStarts);
aPointTable[30].eQuality := F_IiotQuality(xValid := TRUE, iNe107 := TO_INT(GVL_Devices.fbP103.stSts.stCommon.eNe107));
aPointTable[31].lrValue := UINT_TO_LREAL(GVL_Devices.fbP103.stSts.uiStartsLastHour);
aPointTable[31].eQuality := F_IiotQuality(xValid := TRUE, iNe107 := TO_INT(GVL_Devices.fbP103.stSts.stCommon.eNe107));
aPointTable[32].lrValue := REAL_TO_LREAL(GVL_Devices.fbP103.stSts.rRunTimeMaint_h);
aPointTable[32].eQuality := F_IiotQuality(xValid := TRUE, iNe107 := TO_INT(GVL_Devices.fbP103.stSts.stCommon.eNe107));
aPointTable[33].lrValue := UDINT_TO_LREAL(GVL_Devices.fbP103.stSts.udiStartsMaint);
aPointTable[33].eQuality := F_IiotQuality(xValid := TRUE, iNe107 := TO_INT(GVL_Devices.fbP103.stSts.stCommon.eNe107));
aPointTable[34].lrValue := UINT_TO_LREAL(GVL_IO.uiP103_FCODE);
aPointTable[34].eQuality := F_IiotQuality(xValid := TRUE, iNe107 := TO_INT(GVL_Devices.fbP103.stSts.stCommon.eNe107));
IF (GVL_Devices.fbP103.stSts.stCommon.wFault AND PL.GVL_Const.MOT_FLT_COMM_LOSS) <> 0
   OR (GVL_Devices.fbP103.stSts.stCommon.wWarning AND PL.GVL_Const.MOT_WRN_COMM_LOSS) <> 0 THEN
    aPointTable[34].eQuality := E_IiotQuality.Bad;
END_IF
aPointTable[35].lrValue := INT_TO_LREAL(TO_INT(GVL_Devices.fbP103.stSts.stCommon.eMode));
aPointTable[35].eQuality := F_IiotQuality(xValid := TRUE, iNe107 := TO_INT(GVL_Devices.fbP103.stSts.stCommon.eNe107));
aPointTable[36].lrValue := INT_TO_LREAL(TO_INT(GVL_Devices.fbP103.stSts.stCommon.eNe107));
aPointTable[36].eQuality := F_IiotQuality(xValid := TRUE, iNe107 := TO_INT(GVL_Devices.fbP103.stSts.stCommon.eNe107));
aPointTable[37].lrValue := BOOL_TO_LREAL(GVL_Devices.fbV1.xRunning);
aPointTable[37].eQuality := F_IiotQuality(xValid := TRUE, iNe107 := TO_INT(GVL_Devices.fbV1.stSts.stCommon.eNe107));
aPointTable[38].lrValue := INT_TO_LREAL(TO_INT(GVL_Devices.fbV1.stSts.eState));
aPointTable[38].eQuality := F_IiotQuality(xValid := TRUE, iNe107 := TO_INT(GVL_Devices.fbV1.stSts.stCommon.eNe107));
aPointTable[39].lrValue := REAL_TO_LREAL(GVL_Devices.fbV1.stSts.rRunTime_h);
aPointTable[39].eQuality := F_IiotQuality(xValid := TRUE, iNe107 := TO_INT(GVL_Devices.fbV1.stSts.stCommon.eNe107));
aPointTable[40].lrValue := UDINT_TO_LREAL(GVL_Devices.fbV1.stSts.udiStarts);
aPointTable[40].eQuality := F_IiotQuality(xValid := TRUE, iNe107 := TO_INT(GVL_Devices.fbV1.stSts.stCommon.eNe107));
aPointTable[41].lrValue := UINT_TO_LREAL(GVL_Devices.fbV1.stSts.uiStartsLastHour);
aPointTable[41].eQuality := F_IiotQuality(xValid := TRUE, iNe107 := TO_INT(GVL_Devices.fbV1.stSts.stCommon.eNe107));
aPointTable[42].lrValue := REAL_TO_LREAL(GVL_Devices.fbV1.stSts.rRunTimeMaint_h);
aPointTable[42].eQuality := F_IiotQuality(xValid := TRUE, iNe107 := TO_INT(GVL_Devices.fbV1.stSts.stCommon.eNe107));
aPointTable[43].lrValue := UDINT_TO_LREAL(GVL_Devices.fbV1.stSts.udiStartsMaint);
aPointTable[43].eQuality := F_IiotQuality(xValid := TRUE, iNe107 := TO_INT(GVL_Devices.fbV1.stSts.stCommon.eNe107));
aPointTable[44].lrValue := INT_TO_LREAL(TO_INT(GVL_Devices.fbV1.stSts.stCommon.eMode));
aPointTable[44].eQuality := F_IiotQuality(xValid := TRUE, iNe107 := TO_INT(GVL_Devices.fbV1.stSts.stCommon.eNe107));
aPointTable[45].lrValue := INT_TO_LREAL(TO_INT(GVL_Devices.fbV1.stSts.stCommon.eNe107));
aPointTable[45].eQuality := F_IiotQuality(xValid := TRUE, iNe107 := TO_INT(GVL_Devices.fbV1.stSts.stCommon.eNe107));
aPointTable[46].lrValue := REAL_TO_LREAL(GVL_Devices.fbLT101.stSts.rValue_eu);
aPointTable[46].eQuality := F_IiotQuality(xValid := GVL_Devices.fbLT101.xValid,
    iNe107 := TO_INT(GVL_Devices.fbLT101.stSts.stCommon.eNe107));
aPointTable[47].lrValue := INT_TO_LREAL(TO_INT(GVL_Devices.fbLT101.stSts.stCommon.eMode));
aPointTable[47].eQuality := F_IiotQuality(xValid := GVL_Devices.fbLT101.xValid,
    iNe107 := TO_INT(GVL_Devices.fbLT101.stSts.stCommon.eNe107));
aPointTable[48].lrValue := INT_TO_LREAL(TO_INT(GVL_Devices.fbLT101.stSts.stCommon.eNe107));
aPointTable[48].eQuality := F_IiotQuality(xValid := GVL_Devices.fbLT101.xValid,
    iNe107 := TO_INT(GVL_Devices.fbLT101.stSts.stCommon.eNe107));
aPointTable[49].lrValue := BOOL_TO_LREAL(GVL_Devices.fbLS102.xValue);
aPointTable[49].eQuality := F_IiotQuality(xValid := GVL_Devices.fbLS102.xValid,
    iNe107 := TO_INT(GVL_Devices.fbLS102.stSts.stCommon.eNe107));
aPointTable[50].lrValue := INT_TO_LREAL(TO_INT(GVL_Devices.fbLS102.stSts.stCommon.eMode));
aPointTable[50].eQuality := F_IiotQuality(xValid := GVL_Devices.fbLS102.xValid,
    iNe107 := TO_INT(GVL_Devices.fbLS102.stSts.stCommon.eNe107));
aPointTable[51].lrValue := INT_TO_LREAL(TO_INT(GVL_Devices.fbLS102.stSts.stCommon.eNe107));
aPointTable[51].eQuality := F_IiotQuality(xValid := GVL_Devices.fbLS102.xValid,
    iNe107 := TO_INT(GVL_Devices.fbLS102.stSts.stCommon.eNe107));
aPointTable[52].lrValue := BOOL_TO_LREAL(GVL_Devices.fbLS103.xValue);
aPointTable[52].eQuality := F_IiotQuality(xValid := GVL_Devices.fbLS103.xValid,
    iNe107 := TO_INT(GVL_Devices.fbLS103.stSts.stCommon.eNe107));
aPointTable[53].lrValue := INT_TO_LREAL(TO_INT(GVL_Devices.fbLS103.stSts.stCommon.eMode));
aPointTable[53].eQuality := F_IiotQuality(xValid := GVL_Devices.fbLS103.xValid,
    iNe107 := TO_INT(GVL_Devices.fbLS103.stSts.stCommon.eNe107));
aPointTable[54].lrValue := INT_TO_LREAL(TO_INT(GVL_Devices.fbLS103.stSts.stCommon.eNe107));
aPointTable[54].eQuality := F_IiotQuality(xValid := GVL_Devices.fbLS103.xValid,
    iNe107 := TO_INT(GVL_Devices.fbLS103.stSts.stCommon.eNe107));
aPointTable[55].lrValue := REAL_TO_LREAL(GVL_Devices.fbIT111.stSts.rValue_eu);
aPointTable[55].eQuality := F_IiotQuality(xValid := GVL_Devices.fbIT111.xValid,
    iNe107 := TO_INT(GVL_Devices.fbIT111.stSts.stCommon.eNe107));
aPointTable[56].lrValue := INT_TO_LREAL(TO_INT(GVL_Devices.fbIT111.stSts.stCommon.eMode));
aPointTable[56].eQuality := F_IiotQuality(xValid := GVL_Devices.fbIT111.xValid,
    iNe107 := TO_INT(GVL_Devices.fbIT111.stSts.stCommon.eNe107));
aPointTable[57].lrValue := INT_TO_LREAL(TO_INT(GVL_Devices.fbIT111.stSts.stCommon.eNe107));
aPointTable[57].eQuality := F_IiotQuality(xValid := GVL_Devices.fbIT111.xValid,
    iNe107 := TO_INT(GVL_Devices.fbIT111.stSts.stCommon.eNe107));
aPointTable[58].lrValue := BOOL_TO_LREAL(GVL_Devices.fbTS112.xValue);
aPointTable[58].eQuality := F_IiotQuality(xValid := GVL_Devices.fbTS112.xValid,
    iNe107 := TO_INT(GVL_Devices.fbTS112.stSts.stCommon.eNe107));
aPointTable[59].lrValue := INT_TO_LREAL(TO_INT(GVL_Devices.fbTS112.stSts.stCommon.eMode));
aPointTable[59].eQuality := F_IiotQuality(xValid := GVL_Devices.fbTS112.xValid,
    iNe107 := TO_INT(GVL_Devices.fbTS112.stSts.stCommon.eNe107));
aPointTable[60].lrValue := INT_TO_LREAL(TO_INT(GVL_Devices.fbTS112.stSts.stCommon.eNe107));
aPointTable[60].eQuality := F_IiotQuality(xValid := GVL_Devices.fbTS112.xValid,
    iNe107 := TO_INT(GVL_Devices.fbTS112.stSts.stCommon.eNe107));
aPointTable[61].lrValue := BOOL_TO_LREAL(GVL_Devices.fbMS113.xValue);
aPointTable[61].eQuality := F_IiotQuality(xValid := GVL_Devices.fbMS113.xValid,
    iNe107 := TO_INT(GVL_Devices.fbMS113.stSts.stCommon.eNe107));
aPointTable[62].lrValue := INT_TO_LREAL(TO_INT(GVL_Devices.fbMS113.stSts.stCommon.eMode));
aPointTable[62].eQuality := F_IiotQuality(xValid := GVL_Devices.fbMS113.xValid,
    iNe107 := TO_INT(GVL_Devices.fbMS113.stSts.stCommon.eNe107));
aPointTable[63].lrValue := INT_TO_LREAL(TO_INT(GVL_Devices.fbMS113.stSts.stCommon.eNe107));
aPointTable[63].eQuality := F_IiotQuality(xValid := GVL_Devices.fbMS113.xValid,
    iNe107 := TO_INT(GVL_Devices.fbMS113.stSts.stCommon.eNe107));
aPointTable[64].lrValue := REAL_TO_LREAL(GVL_Devices.fbIT121.stSts.rValue_eu);
aPointTable[64].eQuality := F_IiotQuality(xValid := GVL_Devices.fbIT121.xValid,
    iNe107 := TO_INT(GVL_Devices.fbIT121.stSts.stCommon.eNe107));
aPointTable[65].lrValue := INT_TO_LREAL(TO_INT(GVL_Devices.fbIT121.stSts.stCommon.eMode));
aPointTable[65].eQuality := F_IiotQuality(xValid := GVL_Devices.fbIT121.xValid,
    iNe107 := TO_INT(GVL_Devices.fbIT121.stSts.stCommon.eNe107));
aPointTable[66].lrValue := INT_TO_LREAL(TO_INT(GVL_Devices.fbIT121.stSts.stCommon.eNe107));
aPointTable[66].eQuality := F_IiotQuality(xValid := GVL_Devices.fbIT121.xValid,
    iNe107 := TO_INT(GVL_Devices.fbIT121.stSts.stCommon.eNe107));
aPointTable[67].lrValue := BOOL_TO_LREAL(GVL_Devices.fbTS122.xValue);
aPointTable[67].eQuality := F_IiotQuality(xValid := GVL_Devices.fbTS122.xValid,
    iNe107 := TO_INT(GVL_Devices.fbTS122.stSts.stCommon.eNe107));
aPointTable[68].lrValue := INT_TO_LREAL(TO_INT(GVL_Devices.fbTS122.stSts.stCommon.eMode));
aPointTable[68].eQuality := F_IiotQuality(xValid := GVL_Devices.fbTS122.xValid,
    iNe107 := TO_INT(GVL_Devices.fbTS122.stSts.stCommon.eNe107));
aPointTable[69].lrValue := INT_TO_LREAL(TO_INT(GVL_Devices.fbTS122.stSts.stCommon.eNe107));
aPointTable[69].eQuality := F_IiotQuality(xValid := GVL_Devices.fbTS122.xValid,
    iNe107 := TO_INT(GVL_Devices.fbTS122.stSts.stCommon.eNe107));
aPointTable[70].lrValue := BOOL_TO_LREAL(GVL_Devices.fbMS123.xValue);
aPointTable[70].eQuality := F_IiotQuality(xValid := GVL_Devices.fbMS123.xValid,
    iNe107 := TO_INT(GVL_Devices.fbMS123.stSts.stCommon.eNe107));
aPointTable[71].lrValue := INT_TO_LREAL(TO_INT(GVL_Devices.fbMS123.stSts.stCommon.eMode));
aPointTable[71].eQuality := F_IiotQuality(xValid := GVL_Devices.fbMS123.xValid,
    iNe107 := TO_INT(GVL_Devices.fbMS123.stSts.stCommon.eNe107));
aPointTable[72].lrValue := INT_TO_LREAL(TO_INT(GVL_Devices.fbMS123.stSts.stCommon.eNe107));
aPointTable[72].eQuality := F_IiotQuality(xValid := GVL_Devices.fbMS123.xValid,
    iNe107 := TO_INT(GVL_Devices.fbMS123.stSts.stCommon.eNe107));
aPointTable[73].lrValue := REAL_TO_LREAL(GVL_Devices.fbIT131.stSts.rValue_eu);
aPointTable[73].eQuality := F_IiotQuality(xValid := GVL_Devices.fbIT131.xValid,
    iNe107 := TO_INT(GVL_Devices.fbIT131.stSts.stCommon.eNe107));
aPointTable[74].lrValue := INT_TO_LREAL(TO_INT(GVL_Devices.fbIT131.stSts.stCommon.eMode));
aPointTable[74].eQuality := F_IiotQuality(xValid := GVL_Devices.fbIT131.xValid,
    iNe107 := TO_INT(GVL_Devices.fbIT131.stSts.stCommon.eNe107));
aPointTable[75].lrValue := INT_TO_LREAL(TO_INT(GVL_Devices.fbIT131.stSts.stCommon.eNe107));
aPointTable[75].eQuality := F_IiotQuality(xValid := GVL_Devices.fbIT131.xValid,
    iNe107 := TO_INT(GVL_Devices.fbIT131.stSts.stCommon.eNe107));
aPointTable[76].lrValue := BOOL_TO_LREAL(GVL_Devices.fbTS132.xValue);
aPointTable[76].eQuality := F_IiotQuality(xValid := GVL_Devices.fbTS132.xValid,
    iNe107 := TO_INT(GVL_Devices.fbTS132.stSts.stCommon.eNe107));
aPointTable[77].lrValue := INT_TO_LREAL(TO_INT(GVL_Devices.fbTS132.stSts.stCommon.eMode));
aPointTable[77].eQuality := F_IiotQuality(xValid := GVL_Devices.fbTS132.xValid,
    iNe107 := TO_INT(GVL_Devices.fbTS132.stSts.stCommon.eNe107));
aPointTable[78].lrValue := INT_TO_LREAL(TO_INT(GVL_Devices.fbTS132.stSts.stCommon.eNe107));
aPointTable[78].eQuality := F_IiotQuality(xValid := GVL_Devices.fbTS132.xValid,
    iNe107 := TO_INT(GVL_Devices.fbTS132.stSts.stCommon.eNe107));
aPointTable[79].lrValue := BOOL_TO_LREAL(GVL_Devices.fbMS133.xValue);
aPointTable[79].eQuality := F_IiotQuality(xValid := GVL_Devices.fbMS133.xValid,
    iNe107 := TO_INT(GVL_Devices.fbMS133.stSts.stCommon.eNe107));
aPointTable[80].lrValue := INT_TO_LREAL(TO_INT(GVL_Devices.fbMS133.stSts.stCommon.eMode));
aPointTable[80].eQuality := F_IiotQuality(xValid := GVL_Devices.fbMS133.xValid,
    iNe107 := TO_INT(GVL_Devices.fbMS133.stSts.stCommon.eNe107));
aPointTable[81].lrValue := INT_TO_LREAL(TO_INT(GVL_Devices.fbMS133.stSts.stCommon.eNe107));
aPointTable[81].eQuality := F_IiotQuality(xValid := GVL_Devices.fbMS133.xValid,
    iNe107 := TO_INT(GVL_Devices.fbMS133.stSts.stCommon.eNe107));
aPointTable[82].lrValue := REAL_TO_LREAL(GVL_Devices.fbPT201.stSts.rValue_eu);
aPointTable[82].eQuality := F_IiotQuality(xValid := GVL_Devices.fbPT201.xValid,
    iNe107 := TO_INT(GVL_Devices.fbPT201.stSts.stCommon.eNe107));
aPointTable[83].lrValue := INT_TO_LREAL(TO_INT(GVL_Devices.fbPT201.stSts.stCommon.eMode));
aPointTable[83].eQuality := F_IiotQuality(xValid := GVL_Devices.fbPT201.xValid,
    iNe107 := TO_INT(GVL_Devices.fbPT201.stSts.stCommon.eNe107));
aPointTable[84].lrValue := INT_TO_LREAL(TO_INT(GVL_Devices.fbPT201.stSts.stCommon.eNe107));
aPointTable[84].eQuality := F_IiotQuality(xValid := GVL_Devices.fbPT201.xValid,
    iNe107 := TO_INT(GVL_Devices.fbPT201.stSts.stCommon.eNe107));
aPointTable[85].lrValue := REAL_TO_LREAL(GVL_Devices.fbFT202.stSts.rValue_eu);
aPointTable[85].eQuality := F_IiotQuality(xValid := GVL_Devices.fbFT202.xValid,
    iNe107 := TO_INT(GVL_Devices.fbFT202.stSts.stCommon.eNe107));
aPointTable[86].lrValue := INT_TO_LREAL(TO_INT(GVL_Devices.fbFT202.stSts.stCommon.eMode));
aPointTable[86].eQuality := F_IiotQuality(xValid := GVL_Devices.fbFT202.xValid,
    iNe107 := TO_INT(GVL_Devices.fbFT202.stSts.stCommon.eNe107));
aPointTable[87].lrValue := INT_TO_LREAL(TO_INT(GVL_Devices.fbFT202.stSts.stCommon.eNe107));
aPointTable[87].eQuality := F_IiotQuality(xValid := GVL_Devices.fbFT202.xValid,
    iNe107 := TO_INT(GVL_Devices.fbFT202.stSts.stCommon.eNe107));
aPointTable[88].lrValue := BOOL_TO_LREAL(GVL_Devices.fbLS203.xValue);
aPointTable[88].eQuality := F_IiotQuality(xValid := GVL_Devices.fbLS203.xValid,
    iNe107 := TO_INT(GVL_Devices.fbLS203.stSts.stCommon.eNe107));
aPointTable[89].lrValue := INT_TO_LREAL(TO_INT(GVL_Devices.fbLS203.stSts.stCommon.eMode));
aPointTable[89].eQuality := F_IiotQuality(xValid := GVL_Devices.fbLS203.xValid,
    iNe107 := TO_INT(GVL_Devices.fbLS203.stSts.stCommon.eNe107));
aPointTable[90].lrValue := INT_TO_LREAL(TO_INT(GVL_Devices.fbLS203.stSts.stCommon.eNe107));
aPointTable[90].eQuality := F_IiotQuality(xValid := GVL_Devices.fbLS203.xValid,
    iNe107 := TO_INT(GVL_Devices.fbLS203.stSts.stCommon.eNe107));
aPointTable[91].lrValue := BOOL_TO_LREAL(GVL_Devices.fbES301.xValue);
aPointTable[91].eQuality := F_IiotQuality(xValid := GVL_Devices.fbES301.xValid,
    iNe107 := TO_INT(GVL_Devices.fbES301.stSts.stCommon.eNe107));
aPointTable[92].lrValue := INT_TO_LREAL(TO_INT(GVL_Devices.fbES301.stSts.stCommon.eMode));
aPointTable[92].eQuality := F_IiotQuality(xValid := GVL_Devices.fbES301.xValid,
    iNe107 := TO_INT(GVL_Devices.fbES301.stSts.stCommon.eNe107));
aPointTable[93].lrValue := INT_TO_LREAL(TO_INT(GVL_Devices.fbES301.stSts.stCommon.eNe107));
aPointTable[93].eQuality := F_IiotQuality(xValid := GVL_Devices.fbES301.xValid,
    iNe107 := TO_INT(GVL_Devices.fbES301.stSts.stCommon.eNe107));
aPointTable[94].lrValue := BOOL_TO_LREAL(GVL_Devices.fbYS302.xValue);
aPointTable[94].eQuality := F_IiotQuality(xValid := GVL_Devices.fbYS302.xValid,
    iNe107 := TO_INT(GVL_Devices.fbYS302.stSts.stCommon.eNe107));
aPointTable[95].lrValue := INT_TO_LREAL(TO_INT(GVL_Devices.fbYS302.stSts.stCommon.eMode));
aPointTable[95].eQuality := F_IiotQuality(xValid := GVL_Devices.fbYS302.xValid,
    iNe107 := TO_INT(GVL_Devices.fbYS302.stSts.stCommon.eNe107));
aPointTable[96].lrValue := INT_TO_LREAL(TO_INT(GVL_Devices.fbYS302.stSts.stCommon.eNe107));
aPointTable[96].eQuality := F_IiotQuality(xValid := GVL_Devices.fbYS302.xValid,
    iNe107 := TO_INT(GVL_Devices.fbYS302.stSts.stCommon.eNe107));
aPointTable[97].lrValue := BOOL_TO_LREAL(GVL_Devices.fbYS303.xValue);
aPointTable[97].eQuality := F_IiotQuality(xValid := GVL_Devices.fbYS303.xValid,
    iNe107 := TO_INT(GVL_Devices.fbYS303.stSts.stCommon.eNe107));
aPointTable[98].lrValue := INT_TO_LREAL(TO_INT(GVL_Devices.fbYS303.stSts.stCommon.eMode));
aPointTable[98].eQuality := F_IiotQuality(xValid := GVL_Devices.fbYS303.xValid,
    iNe107 := TO_INT(GVL_Devices.fbYS303.stSts.stCommon.eNe107));
aPointTable[99].lrValue := INT_TO_LREAL(TO_INT(GVL_Devices.fbYS303.stSts.stCommon.eNe107));
aPointTable[99].eQuality := F_IiotQuality(xValid := GVL_Devices.fbYS303.xValid,
    iNe107 := TO_INT(GVL_Devices.fbYS303.stSts.stCommon.eNe107));
aPointTable[100].lrValue := REAL_TO_LREAL(GVL_Devices.fbAT401.stSts.rValue_eu);
aPointTable[100].eQuality := F_IiotQuality(xValid := GVL_Devices.fbAT401.xValid,
    iNe107 := TO_INT(GVL_Devices.fbAT401.stSts.stCommon.eNe107));
aPointTable[101].lrValue := INT_TO_LREAL(TO_INT(GVL_Devices.fbAT401.stSts.stCommon.eMode));
aPointTable[101].eQuality := F_IiotQuality(xValid := GVL_Devices.fbAT401.xValid,
    iNe107 := TO_INT(GVL_Devices.fbAT401.stSts.stCommon.eNe107));
aPointTable[102].lrValue := INT_TO_LREAL(TO_INT(GVL_Devices.fbAT401.stSts.stCommon.eNe107));
aPointTable[102].eQuality := F_IiotQuality(xValid := GVL_Devices.fbAT401.xValid,
    iNe107 := TO_INT(GVL_Devices.fbAT401.stSts.stCommon.eNe107));
aPointTable[103].lrValue := REAL_TO_LREAL(GVL_Devices.fbAT402.stSts.rValue_eu);
aPointTable[103].eQuality := F_IiotQuality(xValid := GVL_Devices.fbAT402.xValid,
    iNe107 := TO_INT(GVL_Devices.fbAT402.stSts.stCommon.eNe107));
aPointTable[104].lrValue := INT_TO_LREAL(TO_INT(GVL_Devices.fbAT402.stSts.stCommon.eMode));
aPointTable[104].eQuality := F_IiotQuality(xValid := GVL_Devices.fbAT402.xValid,
    iNe107 := TO_INT(GVL_Devices.fbAT402.stSts.stCommon.eNe107));
aPointTable[105].lrValue := INT_TO_LREAL(TO_INT(GVL_Devices.fbAT402.stSts.stCommon.eNe107));
aPointTable[105].eQuality := F_IiotQuality(xValid := GVL_Devices.fbAT402.xValid,
    iNe107 := TO_INT(GVL_Devices.fbAT402.stSts.stCommon.eNe107));
aPointTable[106].lrValue := REAL_TO_LREAL(GVL_Devices.fbTT403.stSts.rValue_eu);
aPointTable[106].eQuality := F_IiotQuality(xValid := GVL_Devices.fbTT403.xValid,
    iNe107 := TO_INT(GVL_Devices.fbTT403.stSts.stCommon.eNe107));
aPointTable[107].lrValue := INT_TO_LREAL(TO_INT(GVL_Devices.fbTT403.stSts.stCommon.eMode));
aPointTable[107].eQuality := F_IiotQuality(xValid := GVL_Devices.fbTT403.xValid,
    iNe107 := TO_INT(GVL_Devices.fbTT403.stSts.stCommon.eNe107));
aPointTable[108].lrValue := INT_TO_LREAL(TO_INT(GVL_Devices.fbTT403.stSts.stCommon.eNe107));
aPointTable[108].eQuality := F_IiotQuality(xValid := GVL_Devices.fbTT403.xValid,
    iNe107 := TO_INT(GVL_Devices.fbTT403.stSts.stCommon.eNe107));
aPointTable[109].lrValue := BOOL_TO_LREAL(GVL_Devices.fbZS404.xValue);
aPointTable[109].eQuality := F_IiotQuality(xValid := GVL_Devices.fbZS404.xValid,
    iNe107 := TO_INT(GVL_Devices.fbZS404.stSts.stCommon.eNe107));
aPointTable[110].lrValue := INT_TO_LREAL(TO_INT(GVL_Devices.fbZS404.stSts.stCommon.eMode));
aPointTable[110].eQuality := F_IiotQuality(xValid := GVL_Devices.fbZS404.xValid,
    iNe107 := TO_INT(GVL_Devices.fbZS404.stSts.stCommon.eNe107));
aPointTable[111].lrValue := INT_TO_LREAL(TO_INT(GVL_Devices.fbZS404.stSts.stCommon.eNe107));
aPointTable[111].eQuality := F_IiotQuality(xValid := GVL_Devices.fbZS404.xValid,
    iNe107 := TO_INT(GVL_Devices.fbZS404.stSts.stCommon.eNe107));
aPointTable[112].lrValue := BOOL_TO_LREAL(GVL_Devices.fbYS405.xValue);
aPointTable[112].eQuality := F_IiotQuality(xValid := GVL_Devices.fbYS405.xValid,
    iNe107 := TO_INT(GVL_Devices.fbYS405.stSts.stCommon.eNe107));
aPointTable[113].lrValue := INT_TO_LREAL(TO_INT(GVL_Devices.fbYS405.stSts.stCommon.eMode));
aPointTable[113].eQuality := F_IiotQuality(xValid := GVL_Devices.fbYS405.xValid,
    iNe107 := TO_INT(GVL_Devices.fbYS405.stSts.stCommon.eNe107));
aPointTable[114].lrValue := INT_TO_LREAL(TO_INT(GVL_Devices.fbYS405.stSts.stCommon.eNe107));
aPointTable[114].eQuality := F_IiotQuality(xValid := GVL_Devices.fbYS405.xValid,
    iNe107 := TO_INT(GVL_Devices.fbYS405.stSts.stCommon.eNe107));
aPointTable[115].lrValue := BOOL_TO_LREAL(NOT GVL_IO.xK1);
aPointTable[115].eQuality := E_IiotQuality.Good;
aPointTable[116].lrValue := INT_TO_LREAL(TO_INT(GVL_Station.stStationSts.eMode));
aPointTable[116].eQuality := E_IiotQuality.Good;
aPointTable[117].lrValue := INT_TO_LREAL(TO_INT(GVL_Station.stStationSts.eMethod));
aPointTable[117].eQuality := E_IiotQuality.Good;
aPointTable[118].lrValue := INT_TO_LREAL(TO_INT(GVL_Station.stStationSts.eControlAct));
aPointTable[118].eQuality := E_IiotQuality.Good;
aPointTable[119].lrValue := INT_TO_LREAL(TO_INT(GVL_Station.stStationSts.eNe107));
aPointTable[119].eQuality := E_IiotQuality.Good;
aPointTable[120].lrValue := WORD_TO_LREAL(GVL_Station.stStationSts.wState);
aPointTable[120].eQuality := E_IiotQuality.Good;
aPointTable[121].lrValue := UINT_TO_LREAL(GVL_Station.stStationSts.uiPumpsRequired);
aPointTable[121].eQuality := E_IiotQuality.Good;
aPointTable[122].lrValue := UINT_TO_LREAL(GVL_Station.stStationSts.uiPumpsRunning);
aPointTable[122].eQuality := E_IiotQuality.Good;
aPointTable[123].lrValue := UINT_TO_LREAL(GVL_Station.stStationSts.uiPumpsAvailable);
aPointTable[123].eQuality := E_IiotQuality.Good;
aPointTable[124].lrValue := UINT_TO_LREAL(GVL_Station.stStationSts.uiLeadPump);
aPointTable[124].eQuality := E_IiotQuality.Good;
aPointTable[125].lrValue := UINT_TO_LREAL(GVL_Station.stStationSts.uiSeqRemain_s);
aPointTable[125].eQuality := E_IiotQuality.Good;
aPointTable[126].lrValue := REAL_TO_LREAL(GVL_Station.stStationSts.rLevel_m);
aPointTable[126].eQuality := E_IiotQuality.Good;
aPointTable[127].lrValue := REAL_TO_LREAL(GVL_Station.stStationSts.rLevelSp_m);
aPointTable[127].eQuality := E_IiotQuality.Good;
aPointTable[128].lrValue := REAL_TO_LREAL(GVL_Station.stStationSts.rSpeedSp_pct);
aPointTable[128].eQuality := E_IiotQuality.Good;
aPointTable[129].lrValue := REAL_TO_LREAL(GVL_Station.fbLIC101.stSts.rPv_eu);
aPointTable[129].eQuality := F_IiotQuality(xValid := TRUE,
    iNe107 := TO_INT(GVL_Station.fbLIC101.stSts.stCommon.eNe107));
aPointTable[130].lrValue := REAL_TO_LREAL(GVL_Station.fbLIC101.stSts.rSp_eu);
aPointTable[130].eQuality := F_IiotQuality(xValid := TRUE,
    iNe107 := TO_INT(GVL_Station.fbLIC101.stSts.stCommon.eNe107));
aPointTable[131].lrValue := REAL_TO_LREAL(GVL_Station.fbLIC101.stSts.rOut_pct);
aPointTable[131].eQuality := F_IiotQuality(xValid := TRUE,
    iNe107 := TO_INT(GVL_Station.fbLIC101.stSts.stCommon.eNe107));
aPointTable[132].lrValue := INT_TO_LREAL(TO_INT(GVL_Station.fbLIC101.stSts.stCommon.eMode));
aPointTable[132].eQuality := F_IiotQuality(xValid := TRUE,
    iNe107 := TO_INT(GVL_Station.fbLIC101.stSts.stCommon.eNe107));
aPointTable[133].lrValue := INT_TO_LREAL(TO_INT(GVL_Station.fbLIC101.stSts.stCommon.eNe107));
aPointTable[133].eQuality := F_IiotQuality(xValid := TRUE,
    iNe107 := TO_INT(GVL_Station.fbLIC101.stSts.stCommon.eNe107));
